(* IEC 61131-3 sources: sis-interlock-demo/pytests/golden/mini/src/POUs/Generated/F_SisIoNormal, 1 file *)

(* ---- F_SisIoNormal.decl.st ---- *)
// AUTO-GENERATED by cemgen 1.0.0 — не редактировать: правьте матрицу и запустите
//   python -m cemgen generate <файл матрицы .csv или .xlsx>
// Матрица: TEST-U301-CEM, объект U-301, ревизия 1 от 2026-10-16, SHA-256 сетки 9067fda96ae55e67
// Назначение: нормальное состояние образа ввода-вывода: все каналы в норме и достоверны, контроль
//             линии исправен, ключи и кнопка не нажаты; выходы xQ* не трогает. Для демо без
//             ввода-вывода и тестов. Возвращает TRUE.
// Автор:      pytest; код — генератор cemgen
// Версия:     1.0.0
// Документ:   docs/DESIGN.md, раздел «10. Генератор cemgen»; docs/cause_effect_matrix.md
// ВНИМАНИЕ:   код демонстрационный и не предназначен для систем безопасности. Реальная ПАЗ требует
//             определения SIL, сертифицированных аппаратных и программных средств и валидации по
//             ГОСТ Р МЭК 61511.
FUNCTION F_SisIoNormal : BOOL
VAR_IN_OUT
    stIo : ST_SisIo;   // образ ввода-вывода
END_VAR
